(* IEC 61131-3 sources: avi-aoi-management/server/services/programming/iec61131/golden-st/invalid, 40 files *)

(* ---- i34-fb-member-not-declared.st ---- *)
FUNCTION_BLOCK FB_Motor
VAR_INPUT
    Run : BOOL;
END_VAR
VAR_OUTPUT
    Running : BOOL;
END_VAR
Running := Run;
END_FUNCTION_BLOCK

PROGRAM UseMotor
VAR
    M1   : FB_Motor;
    Lamp : BOOL;
END_VAR
M1(Run := TRUE);
Lamp := M1.IsRunning;
END_PROGRAM

(* ---- i01-probe-garbage.st ---- *)
PROGRAM P
VAR a : BOOL END_VAR
a := TRUE
b = FALSE;;
FOO BAR BAZ (((
MOVEABS(10,20)
END_PROGRAM

(* ---- i02-missing-semicolon.st ---- *)
PROGRAM MissingSemi
VAR
    Start : BOOL;
    Motor : BOOL;
    Lamp  : BOOL;
END_VAR

Motor := Start
Lamp := Motor;

END_PROGRAM

(* ---- i03-if-without-end-if.st ---- *)
PROGRAM NoEndIf
VAR
    Level : INT;
    Pump  : BOOL;
END_VAR

IF Level > 80 THEN
    Pump := FALSE;
ELSE
    Pump := TRUE;

END_PROGRAM

(* ---- i04-ton-member-out.st ---- *)
PROGRAM WrongTimerMember
VAR
    Go   : BOOL;
    Tmr  : TON;
    Lamp : BOOL;
END_VAR

Tmr(IN := Go, PT := T#2s);
Lamp := Tmr.OUT;

END_PROGRAM

(* ---- i05-undeclared-in-expression.st ---- *)
PROGRAM UndeclaredRead
VAR
    Motor : BOOL;
END_VAR

Motor := StartButton AND NOT Motor;

END_PROGRAM

(* ---- i06-undeclared-assignment-target.st ---- *)
PROGRAM UndeclaredWrite
VAR
    Start : BOOL;
END_VAR

ConveyorOn := Start;

END_PROGRAM

(* ---- i07-equals-instead-of-assign.st ---- *)
PROGRAM EqualsAssign
VAR
    Start : BOOL;
    Motor : BOOL;
END_VAR

Motor = Start;

END_PROGRAM

(* ---- i08-double-equals-compare.st ---- *)
PROGRAM DoubleEquals
VAR
    Level : INT;
    Alarm : BOOL;
END_VAR

IF Level == 100 THEN
    Alarm := TRUE;
END_IF;

END_PROGRAM

(* ---- i09-for-without-end-for.st ---- *)
PROGRAM NoEndFor
VAR
    I   : INT;
    Sum : INT;
END_VAR

Sum := 0;
FOR I := 1 TO 10 DO
    Sum := Sum + I;

END_PROGRAM

(* ---- i10-while-missing-do.st ---- *)
PROGRAM WhileNoDo
VAR
    N : INT;
END_VAR

N := 10;
WHILE N > 0
    N := N - 1;
END_WHILE;

END_PROGRAM

(* ---- i11-case-without-end-case.st ---- *)
PROGRAM NoEndCase
VAR
    Step  : INT;
    Valve : BOOL;
END_VAR

CASE Step OF
    0: Valve := FALSE;
    1: Valve := TRUE;

END_PROGRAM

(* ---- i12-repeat-without-until.st ---- *)
PROGRAM RepeatNoUntil
VAR
    K : INT;
END_VAR

REPEAT
    K := K + 1;
END_REPEAT;

END_PROGRAM

(* ---- i13-unterminated-comment.st ---- *)
PROGRAM OpenComment
VAR
    Lamp : BOOL;
END_VAR

(* the lamp follows the door switch
Lamp := TRUE;

END_PROGRAM

(* ---- i14-unterminated-string.st ---- *)
PROGRAM OpenString
VAR
    Msg : STRING;
END_VAR

Msg := 'Line 1 ready;

END_PROGRAM

(* ---- i15-missing-end-var.st ---- *)
PROGRAM NoEndVar
VAR
    Start : BOOL;
    Motor : BOOL;

Motor := Start;

END_PROGRAM

(* ---- i16-missing-end-program.st ---- *)
PROGRAM NoEndProgram
VAR
    Start : BOOL;
    Motor : BOOL;
END_VAR

Motor := Start;

(* ---- i17-ton-bad-input-param.st ---- *)
PROGRAM BadTimerParam
VAR
    Go   : BOOL;
    Tmr  : TON;
    Lamp : BOOL;
END_VAR

Tmr(IN := Go, PRESET := T#2s);
Lamp := Tmr.Q;

END_PROGRAM

(* ---- i18-ctu-member-acc.st ---- *)
PROGRAM AllenBradleyStyle
VAR
    Pulse : BOOL;
    Cnt   : CTU;
    Total : INT;
END_VAR

Cnt(CU := Pulse, R := FALSE, PV := 10);
Total := Cnt.ACC;

END_PROGRAM

(* ---- i19-undeclared-fb-instance.st ---- *)
PROGRAM NoInstance
VAR
    Go   : BOOL;
    Lamp : BOOL;
END_VAR

Timer1(IN := Go, PT := T#1s);
Lamp := Timer1.Q;

END_PROGRAM

(* ---- i20-bad-time-literal.st ---- *)
PROGRAM BadTime
VAR
    Go   : BOOL;
    Tmr  : TON;
END_VAR

Tmr(IN := Go, PT := T#2x);

END_PROGRAM

(* ---- i21-elseif-one-word.st ---- *)
PROGRAM ElseIfWord
VAR
    Level : INT;
    Pump  : BOOL;
    Alarm : BOOL;
END_VAR

IF Level > 90 THEN
    Pump := FALSE;
ELSEIF Level > 95 THEN
    Alarm := TRUE;
END_IF;

END_PROGRAM

(* ---- i22-unbalanced-parenthesis.st ---- *)
PROGRAM OpenParen
VAR
    A : BOOL;
    B : BOOL;
    C : BOOL;
END_VAR

C := (A AND B;

END_PROGRAM

(* ---- i23-markdown-fence-prose.st ---- *)
Here is the Structured Text program you asked for:
```iecst
PROGRAM Conveyor
VAR
    Start : BOOL;
    Motor : BOOL;
END_VAR
Motor := Start;
END_PROGRAM
```

(* ---- i24-statement-outside-pou.st ---- *)
PROGRAM Inside
VAR
    Start : BOOL;
    Motor : BOOL;
END_VAR
Motor := Start;
END_PROGRAM

Motor := FALSE;

(* ---- i25-member-on-bool.st ---- *)
PROGRAM MemberOnBool
VAR
    Start : BOOL;
    Lamp  : BOOL;
END_VAR

Lamp := Start.Q;

END_PROGRAM

(* ---- i26-if-closed-by-end-for.st ---- *)
PROGRAM WrongCloser
VAR
    Level : INT;
    Pump  : BOOL;
END_VAR

IF Level > 80 THEN
    Pump := FALSE;
END_FOR;

END_PROGRAM

(* ---- i27-end-if-only-in-comment.st ---- *)
PROGRAM EndIfInComment
VAR
    Door : BOOL;
    Lamp : BOOL;
END_VAR

IF Door THEN
    Lamp := TRUE;
    (* END_IF *)

END_PROGRAM

(* ---- i28-undeclared-for-counter.st ---- *)
PROGRAM UndeclaredCounter
VAR
    Sum : INT;
END_VAR

Sum := 0;
FOR Idx := 1 TO 10 DO
    Sum := Sum + 1;
END_FOR;

END_PROGRAM

(* ---- i29-duplicate-declaration.st ---- *)
PROGRAM Duplicate
VAR
    Motor : BOOL;
    Speed : INT;
    Motor : BOOL;
END_VAR

Motor := Speed > 0;

END_PROGRAM

(* ---- i30-assign-to-constant.st ---- *)
PROGRAM WriteConstant
VAR CONSTANT
    MAX_SPEED : INT := 1500;
END_VAR
VAR
    Speed : INT;
END_VAR

MAX_SPEED := Speed;

END_PROGRAM

(* ---- i31-c-style-operators.st ---- *)
PROGRAM CStyle
VAR
    A : BOOL;
    B : BOOL;
    C : BOOL;
END_VAR

C := A && B;

END_PROGRAM

(* ---- i32-output-bound-to-undeclared.st ---- *)
PROGRAM UndeclaredOutput
VAR
    Go  : BOOL;
    Tmr : TON;
END_VAR

Tmr(IN := Go, PT := T#1s, Q => DoneFlag);

END_PROGRAM

(* ---- i33-then-missing.st ---- *)
PROGRAM ThenMissing
VAR
    Door : BOOL;
    Lamp : BOOL;
END_VAR

IF Door
    Lamp := TRUE;
END_IF;

END_PROGRAM

(* ---- i35-nested-comment.st ---- *)
PROGRAM NestedComment
VAR
    Lamp : BOOL;
END_VAR

(* disabled for commissioning:
   (* old logic *)
   Lamp := FALSE;
*)
Lamp := TRUE;

END_PROGRAM

(* ---- i36-r-edge-outside-var-input.st ---- *)
PROGRAM EdgeInLocalVar
VAR
    Sensor : BOOL R_EDGE;
    Count  : INT;
END_VAR

IF Sensor THEN
    Count := Count + 1;
END_IF;

END_PROGRAM

(* ---- i37-misspelled-time-function.st ---- *)
PROGRAM MisspelledTimeFn
VAR
    Dwell : TIME := T#2s;
    Total : TIME;
END_VAR

Total := ADD_TIMES(Dwell, T#1s);

END_PROGRAM

(* ---- i38-misspelled-limit.st ---- *)
PROGRAM MisspelledLimit
VAR
    Speed : INT;
    Out   : INT;
END_VAR

Out := LIMT(0, Speed, 100);

END_PROGRAM

(* ---- i39-hallucinated-conversion.st ---- *)
PROGRAM HallucinatedConversion
VAR
    Level : INT;
    Out   : REAL;
END_VAR

Out := FOO_BAR_TO_BAZ_QUX(Level);

END_PROGRAM

(* ---- i40-conversion-to-unknown-type.st ---- *)
PROGRAM ConversionToUnknownType
VAR
    Level : INT;
    Out   : REAL;
END_VAR

Out := INT_TO_FOO(Level);

END_PROGRAM
